(* IEC 61131-3 sources: volt/packages/volt-lsp-iec/test-corpus/pro2193/Device/Plc Logic/Application/09 Misc/Library Manager/CmpCodeMeter, 19 files *)

(* ---- EVTPARAM_CMPCODEMETERLICENSEACTIVATED.dut ---- *)
TYPE EVTPARAM_CMPCODEMETERLICENSEACTIVATED :
STRUCT
	SERIALNO : DWORD;
	PSZUPDATEFILE : POINTER TO STRING;
END_STRUCT
END_TYPE

(* ---- RTS_CMBOXENTRY.dut ---- *)
TYPE RTS_CMBOXENTRY :
STRUCT
	MUSBOXMASK : WORD;
	MULBOXSERIAL : UDINT;
	MFLFICTRL : UDINT;
	MULFIRMCODE : UDINT;
	MUSFIRMACCESSCOUNTER : WORD;
	MUSFIRMITEMREF : WORD;
	MULFIRMUPDATECOUNTER : UDINT;
	MULFIRMPRECISETIME : UDINT;
	MAUSFIRMITEMTEXT : WSTRING(255);
	MULPRODUCTCODE : UDINT;
	MULFEATUREMAP : UDINT;
	MULUNITCOUNTER : UDINT;
	MULLICENSEQUANTITY : UDINT;
	MUSPRODUCTITEMREF : WORD;
END_STRUCT
END_TYPE

(* ---- RTS_CODEMETER_INFO.dut ---- *)
TYPE RTS_CODEMETER_INFO :
STRUCT
	BYMAJORVERSION : BYTE;
	BYMINORVERSION : BYTE;
	WBOXMASK : WORD;
	DWSERIALNUMBER : DWORD;
	WCHIPTYPE : WORD;
	WSILICONREVISION : WORD;
END_STRUCT
END_TYPE

(* ---- EVENTIDS.gvl ---- *)
VAR_GLOBAL
	CMPID_CMPCODEMETER : DWORD := 16#7A;
	EVTPARAMID_CMPCODEMETER_LICENSEACTIVATED : WORD := 16#1;
	EVTVERSION_CMPCODEMETER_LICENSEACTIVATED : WORD := 16#1;
	EVT_CMPCODEMETER_LICENSEACTIVATED : DWORD := (SHL(UINT_TO_DWORD(EVTCLASS_INFO), 16) OR 16#1);
END_VAR

(* ---- CODEMCLOSE.pou ---- *)
FUNCTION CODEMCLOSE : RTS_IEC_RESULT
VAR_INPUT
	HCODEMETER : RTS_IEC_HANDLE;
END_VAR
END_FUNCTION

(* ---- CODEMDECREMENTUNITCOUNTER.pou ---- *)
FUNCTION CODEMDECREMENTUNITCOUNTER : RTS_IEC_RESULT
VAR_INPUT
	HCODEMETER : RTS_IEC_HANDLE;
	UDIUNITCOUNT : UDINT;
END_VAR
END_FUNCTION

(* ---- CODEMDECRYPT.pou ---- *)
FUNCTION CODEMDECRYPT : RTS_IEC_RESULT
VAR_INPUT
	HCODEMETER : RTS_IEC_HANDLE;
	UDIENCRYPTIONCODE : UDINT;
	ULCRC : UDINT;
	PBYDATA : POINTER TO BYTE;
	NDATALEN : __XWORD;
END_VAR
END_FUNCTION

(* ---- CODEMENCRYPT.pou ---- *)
FUNCTION CODEMENCRYPT : RTS_IEC_RESULT
VAR_INPUT
	HCODEMETER : RTS_IEC_HANDLE;
	UDIENCRYPTIONCODE : UDINT;
	PBYDATA : POINTER TO BYTE;
	NDATALEN : __XWORD;
END_VAR
VAR_IN_OUT
	ULCRC : UDINT;
END_VAR
END_FUNCTION

(* ---- CODEMGETCONTENTBYFIRMCODE.pou ---- *)
FUNCTION CODEMGETCONTENTBYFIRMCODE : RTS_IEC_RESULT
VAR_INPUT
	DUIFIRMCODE : UDINT;
	DUIPRODUCTCODE : UDINT;
END_VAR
VAR_IN_OUT
	LICENSEENTRY : RTS_CMBOXENTRY;
END_VAR
END_FUNCTION

(* ---- CODEMGETCONTENTBYFIRMCODE2.pou ---- *)
FUNCTION CODEMGETCONTENTBYFIRMCODE2 : RTS_IEC_RESULT
VAR_INPUT
	DUIFIRMCODE : UDINT;
	DUIPRODUCTCODE : UDINT;
	BRELEASELICENSE : BOOL;
END_VAR
VAR_IN_OUT
	LICENSEENTRY : RTS_CMBOXENTRY;
END_VAR
END_FUNCTION

(* ---- CODEMGETEXPIRATIONTIME.pou ---- *)
FUNCTION CODEMGETEXPIRATIONTIME : RTS_IEC_RESULT
VAR_INPUT
	HCODEMETER : RTS_IEC_HANDLE;
END_VAR
VAR_IN_OUT
	DTEXPIRATION : DATE_AND_TIME;
END_VAR
END_FUNCTION

(* ---- CODEMGETFEATUREMAPBYFIRMCODE.pou ---- *)
FUNCTION CODEMGETFEATUREMAPBYFIRMCODE : UDINT
VAR_INPUT
	DUIFIRMCODE : UDINT;
	DUIPRODUCTCODE : UDINT;
END_VAR
END_FUNCTION

(* ---- CODEMGETFIRST.pou ---- *)
FUNCTION CODEMGETFIRST : RTS_IEC_HANDLE
VAR_IN_OUT
	RESULT : RTS_IEC_RESULT;
END_VAR
END_FUNCTION

(* ---- CODEMGETINFO.pou ---- *)
FUNCTION CODEMGETINFO : RTS_IEC_RESULT
VAR_INPUT
	HCODEMETER : RTS_IEC_HANDLE;
END_VAR
VAR_IN_OUT
	INFO : RTS_CODEMETER_INFO;
END_VAR
END_FUNCTION

(* ---- CODEMGETNAME.pou ---- *)
FUNCTION CODEMGETNAME : RTS_IEC_RESULT
VAR_INPUT
	HCODEMETER : RTS_IEC_HANDLE;
	NLENBYTES : UDINT;
END_VAR
VAR_IN_OUT
	WSTNAME : WSTRING(255);
END_VAR
END_FUNCTION

(* ---- CODEMGETNEXT.pou ---- *)
FUNCTION CODEMGETNEXT : RTS_IEC_HANDLE
VAR_INPUT
	HPREVCODEMETER : RTS_IEC_HANDLE;
END_VAR
VAR_IN_OUT
	RESULT : RTS_IEC_RESULT;
END_VAR
END_FUNCTION

(* ---- CODEMGETQUANTITY.pou ---- *)
FUNCTION CODEMGETQUANTITY : RTS_IEC_RESULT
VAR_INPUT
	HCODEMETER : RTS_IEC_HANDLE;
END_VAR
VAR_IN_OUT
	UDIQUANTITY : UDINT;
END_VAR
END_FUNCTION

(* ---- CODEMGETUNITCOUNTER.pou ---- *)
FUNCTION CODEMGETUNITCOUNTER : RTS_IEC_RESULT
VAR_INPUT
	HCODEMETER : RTS_IEC_HANDLE;
END_VAR
VAR_IN_OUT
	UDIUNITCOUNT : UDINT;
END_VAR
END_FUNCTION

(* ---- CODEMOPEN.pou ---- *)
FUNCTION CODEMOPEN : RTS_IEC_HANDLE
VAR_INPUT
	UDIFIRMCODE : UDINT;
	UDIPRODUCTCODE : UDINT;
	UDIFEATURECODE : UDINT;
END_VAR
VAR_IN_OUT
	RESULT : RTS_IEC_RESULT;
END_VAR
END_FUNCTION
